TYPE "ST_TwoHandOutImm"
VERSION : 0.1
   STRUCT
      LeftPressed : Bool;
      RightPressed : Bool;
      SafeActive : Bool;
      Armed : Bool;
      StartPulse : Bool;
      FieldbusHealthy : Bool;
   END_STRUCT;

END_TYPE

